DATA_BLOCK "DB_ExampleCylinder"
{ S7_Optimized_Access := 'FALSE' }
VERSION : 0.1
NON_RETAIN
   STRUCT
      PLCToComso : Struct
         Test_ProNum : Byte;
         ManStart : Bool;
         AutoStart : Bool;
      END_STRUCT;
      ComsoToPLC : Struct
         Test_NG : Bool;
         Test_OK : Bool;
         Running : Bool;
         Test_Date : Real;
      END_STRUCT;
   END_STRUCT;


BEGIN

END_DATA_BLOCK

